(* IEC 61131-3 sources: trust-platform/examples/OSCAT/cip_wash_state/oop/src, 3 files *)

(* ---- Main.st ---- *)
(* Pattern role: ICipState is the contract boundary for the State example. *)
INTERFACE ICipState
    PROPERTY StateId : INT
    GET
    END_GET
    END_PROPERTY

    METHOD OnEnter
    END_METHOD

    METHOD OnExecute : INT
    VAR_INPUT
        StartCommand : BOOL;
        StepComplete : BOOL;
        ConductivityUs : REAL;
        CausticTempC : REAL;
        FlowOk : BOOL;
        EStopHealthy : BOOL;
    END_VAR
    END_METHOD

    METHOD OnExit
    END_METHOD

    METHOD CanAbort : BOOL
    END_METHOD
END_INTERFACE

(* Pattern role: IdleState is a concrete implementation in the State example. *)
FUNCTION_BLOCK IdleState IMPLEMENTS ICipState
VAR
    Entered : BOOL;
END_VAR

METHOD PUBLIC OnEnter
Entered := TRUE;
END_METHOD

METHOD PUBLIC OnExecute : INT
VAR_INPUT
    StartCommand : BOOL;
    StepComplete : BOOL;
    ConductivityUs : REAL;
    CausticTempC : REAL;
    FlowOk : BOOL;
    EStopHealthy : BOOL;
END_VAR
IF NOT EStopHealthy THEN
    OnExecute := INT#90;
ELSIF StartCommand THEN
    OnExecute := INT#10;
ELSE
    OnExecute := INT#0;
END_IF;
END_METHOD

METHOD PUBLIC OnExit
Entered := FALSE;
END_METHOD

METHOD PUBLIC CanAbort : BOOL
CanAbort := TRUE;
END_METHOD

PUBLIC PROPERTY StateId : INT
GET
    StateId := INT#0;
END_GET
END_PROPERTY
END_FUNCTION_BLOCK

(* Pattern role: PreRinseState is a concrete implementation in the State example. *)
FUNCTION_BLOCK PreRinseState IMPLEMENTS ICipState
METHOD PUBLIC OnEnter
END_METHOD

METHOD PUBLIC OnExecute : INT
VAR_INPUT
    StartCommand : BOOL;
    StepComplete : BOOL;
    ConductivityUs : REAL;
    CausticTempC : REAL;
    FlowOk : BOOL;
    EStopHealthy : BOOL;
END_VAR
IF NOT EStopHealthy OR NOT FlowOk THEN
    OnExecute := INT#90;
ELSIF StepComplete THEN
    OnExecute := INT#20;
ELSE
    OnExecute := INT#10;
END_IF;
END_METHOD

METHOD PUBLIC OnExit
END_METHOD

METHOD PUBLIC CanAbort : BOOL
CanAbort := TRUE;
END_METHOD

PUBLIC PROPERTY StateId : INT
GET
    StateId := INT#10;
END_GET
END_PROPERTY
END_FUNCTION_BLOCK

(* Pattern role: CausticWashState is a concrete implementation in the State example. *)
FUNCTION_BLOCK CausticWashState IMPLEMENTS ICipState
METHOD PUBLIC OnEnter
END_METHOD

METHOD PUBLIC OnExecute : INT
VAR_INPUT
    StartCommand : BOOL;
    StepComplete : BOOL;
    ConductivityUs : REAL;
    CausticTempC : REAL;
    FlowOk : BOOL;
    EStopHealthy : BOOL;
END_VAR
IF NOT EStopHealthy OR NOT FlowOk THEN
    OnExecute := INT#90;
ELSIF CausticTempC < REAL#70.0 THEN
    OnExecute := INT#20;
ELSIF StepComplete THEN
    OnExecute := INT#30;
ELSE
    OnExecute := INT#20;
END_IF;
END_METHOD

METHOD PUBLIC OnExit
END_METHOD

METHOD PUBLIC CanAbort : BOOL
CanAbort := TRUE;
END_METHOD

PUBLIC PROPERTY StateId : INT
GET
    StateId := INT#20;
END_GET
END_PROPERTY
END_FUNCTION_BLOCK

(* Pattern role: IntermediateRinseState is a concrete implementation in the State example. *)
FUNCTION_BLOCK IntermediateRinseState IMPLEMENTS ICipState
METHOD PUBLIC OnEnter
END_METHOD

METHOD PUBLIC OnExecute : INT
VAR_INPUT
    StartCommand : BOOL;
    StepComplete : BOOL;
    ConductivityUs : REAL;
    CausticTempC : REAL;
    FlowOk : BOOL;
    EStopHealthy : BOOL;
END_VAR
IF NOT EStopHealthy OR NOT FlowOk THEN
    OnExecute := INT#90;
ELSIF StepComplete THEN
    OnExecute := INT#40;
ELSE
    OnExecute := INT#30;
END_IF;
END_METHOD

METHOD PUBLIC OnExit
END_METHOD

METHOD PUBLIC CanAbort : BOOL
CanAbort := TRUE;
END_METHOD

PUBLIC PROPERTY StateId : INT
GET
    StateId := INT#30;
END_GET
END_PROPERTY
END_FUNCTION_BLOCK

(* Pattern role: AcidWashState is a concrete implementation in the State example. *)
FUNCTION_BLOCK AcidWashState IMPLEMENTS ICipState
METHOD PUBLIC OnEnter
END_METHOD

METHOD PUBLIC OnExecute : INT
VAR_INPUT
    StartCommand : BOOL;
    StepComplete : BOOL;
    ConductivityUs : REAL;
    CausticTempC : REAL;
    FlowOk : BOOL;
    EStopHealthy : BOOL;
END_VAR
IF NOT EStopHealthy OR NOT FlowOk THEN
    OnExecute := INT#90;
ELSIF StepComplete THEN
    OnExecute := INT#50;
ELSE
    OnExecute := INT#40;
END_IF;
END_METHOD

METHOD PUBLIC OnExit
END_METHOD

METHOD PUBLIC CanAbort : BOOL
CanAbort := TRUE;
END_METHOD

PUBLIC PROPERTY StateId : INT
GET
    StateId := INT#40;
END_GET
END_PROPERTY
END_FUNCTION_BLOCK

(* Pattern role: FinalRinseState is a concrete implementation in the State example. *)
FUNCTION_BLOCK FinalRinseState IMPLEMENTS ICipState
METHOD PUBLIC OnEnter
END_METHOD

METHOD PUBLIC OnExecute : INT
VAR_INPUT
    StartCommand : BOOL;
    StepComplete : BOOL;
    ConductivityUs : REAL;
    CausticTempC : REAL;
    FlowOk : BOOL;
    EStopHealthy : BOOL;
END_VAR
IF NOT EStopHealthy OR NOT FlowOk THEN
    OnExecute := INT#90;
ELSIF ConductivityUs < REAL#50.0 THEN
    OnExecute := INT#100;
ELSE
    OnExecute := INT#50;
END_IF;
END_METHOD

METHOD PUBLIC OnExit
END_METHOD

METHOD PUBLIC CanAbort : BOOL
CanAbort := TRUE;
END_METHOD

PUBLIC PROPERTY StateId : INT
GET
    StateId := INT#50;
END_GET
END_PROPERTY
END_FUNCTION_BLOCK

(* Pattern role: DoneState is a concrete implementation in the State example. *)
FUNCTION_BLOCK DoneState IMPLEMENTS ICipState
METHOD PUBLIC OnEnter
END_METHOD

METHOD PUBLIC OnExecute : INT
VAR_INPUT
    StartCommand : BOOL;
    StepComplete : BOOL;
    ConductivityUs : REAL;
    CausticTempC : REAL;
    FlowOk : BOOL;
    EStopHealthy : BOOL;
END_VAR
OnExecute := INT#100;
END_METHOD

METHOD PUBLIC OnExit
END_METHOD

METHOD PUBLIC CanAbort : BOOL
CanAbort := FALSE;
END_METHOD

PUBLIC PROPERTY StateId : INT
GET
    StateId := INT#100;
END_GET
END_PROPERTY
END_FUNCTION_BLOCK

(* Pattern role: AbortState is a concrete implementation in the State example. *)
FUNCTION_BLOCK AbortState IMPLEMENTS ICipState
METHOD PUBLIC OnEnter
END_METHOD

METHOD PUBLIC OnExecute : INT
VAR_INPUT
    StartCommand : BOOL;
    StepComplete : BOOL;
    ConductivityUs : REAL;
    CausticTempC : REAL;
    FlowOk : BOOL;
    EStopHealthy : BOOL;
END_VAR
OnExecute := INT#90;
END_METHOD

METHOD PUBLIC OnExit
END_METHOD

METHOD PUBLIC CanAbort : BOOL
CanAbort := FALSE;
END_METHOD

PUBLIC PROPERTY StateId : INT
GET
    StateId := INT#90;
END_GET
END_PROPERTY
END_FUNCTION_BLOCK

(* Composition role: CipController owns the collaborating objects used by this State example. *)
FUNCTION_BLOCK CipController
VAR
    Idle : IdleState;
    PreRinse : PreRinseState;
    Caustic : CausticWashState;
    Intermediate : IntermediateRinseState;
    Acid : AcidWashState;
    FinalRinse : FinalRinseState;
    CompleteState : DoneState;
    Abort : AbortState;
    Current : ICipState;
    ConductivityFilter : Pt1Filter;
    CycleCounter : DwordCounter;
    CurrentStateIdValue : INT;
    TransitionCountValue : INT;
    AbortedValue : BOOL;
END_VAR

METHOD PUBLIC Initialize
ConductivityFilter.Initialize();
ConductivityFilter.Configure(TimeConstant := T#1s, Gain := REAL#1.0);
CycleCounter.Initialize();
CycleCounter.Configure(StepSize := DWORD#1, MaxValue := DWORD#16#FFFFFFFF);
Current := Idle;
Current.OnEnter();
CurrentStateIdValue := Current.StateId;
TransitionCountValue := INT#0;
AbortedValue := FALSE;
END_METHOD

METHOD PUBLIC ResolveState : ICipState
VAR_INPUT
    NextId : INT;
END_VAR
IF NextId = INT#10 THEN
    ResolveState := PreRinse;
ELSIF NextId = INT#20 THEN
    ResolveState := Caustic;
ELSIF NextId = INT#30 THEN
    ResolveState := Intermediate;
ELSIF NextId = INT#40 THEN
    ResolveState := Acid;
ELSIF NextId = INT#50 THEN
    ResolveState := FinalRinse;
ELSIF NextId = INT#90 THEN
    ResolveState := Abort;
ELSIF NextId = INT#100 THEN
    ResolveState := CompleteState;
ELSE
    ResolveState := Idle;
END_IF;
END_METHOD

METHOD PUBLIC Update : INT
VAR_INPUT
    StartCommand : BOOL;
    StepComplete : BOOL;
    ConductivityUs : REAL;
    CausticTempC : REAL;
    FlowOk : BOOL;
    EStopHealthy : BOOL;
END_VAR
VAR
    NextId : INT;
END_VAR
(* ConductivityFilter is declared and updated for telemetry/HMI use only.
   FinalRinseState compares against the raw ConductivityUs because the
   PT1 filter time constant (1 s) would otherwise delay the wash-complete
   decision past one scan cycle. A production CIP could drive the state
   from the filtered value with a longer minimum-rinse time. *)
ConductivityFilter.Update(Sample := ConductivityUs);
NextId := Current.OnExecute(StartCommand := StartCommand, StepComplete := StepComplete, ConductivityUs := ConductivityUs, CausticTempC := CausticTempC, FlowOk := FlowOk, EStopHealthy := EStopHealthy);
IF NextId <> Current.StateId THEN
    Current.OnExit();
    Current := ResolveState(NextId := NextId);
    Current.OnEnter();
    CurrentStateIdValue := Current.StateId;
    TransitionCountValue := TransitionCountValue + INT#1;
    IF CurrentStateIdValue = INT#90 THEN
        AbortedValue := TRUE;
    ELSIF CurrentStateIdValue = INT#100 THEN
        CycleCounter.Update(Up := TRUE, Down := FALSE);
    END_IF;
END_IF;
Update := CurrentStateIdValue;
END_METHOD

PUBLIC PROPERTY CurrentStateId : INT
GET
    CurrentStateId := CurrentStateIdValue;
END_GET
END_PROPERTY

PUBLIC PROPERTY TransitionCount : INT
GET
    TransitionCount := TransitionCountValue;
END_GET
END_PROPERTY

PUBLIC PROPERTY CycleCount : DWORD
GET
    CycleCount := CycleCounter.Count;
END_GET
END_PROPERTY

PUBLIC PROPERTY Aborted : BOOL
GET
    Aborted := AbortedValue;
END_GET
END_PROPERTY
END_FUNCTION_BLOCK

(* Scan role: Main wires the example objects and exposes the PLC call path under test. *)
PROGRAM Main
VAR
    Cip : CipController;
    Initialized : BOOL;
    StartCommand : BOOL;
    StepComplete : BOOL;
    EStopHealthy : BOOL;
    FlowOk : BOOL;
    ConductivityRaw : INT;
    CausticTempRaw : INT;
    PumpEnableOut : BOOL;
    DrainValveOut : BOOL;
    AlarmOut : BOOL;
END_VAR

(* Initialize once on cold start; scanning Initialize every cycle would
   reset the state machine to Idle and clear retained counters. *)
IF NOT Initialized THEN
    Cip.Initialize();
    Initialized := TRUE;
END_IF;
Cip.Update(StartCommand := StartCommand, StepComplete := StepComplete, ConductivityUs := INT_TO_REAL(ConductivityRaw), CausticTempC := INT_TO_REAL(CausticTempRaw), FlowOk := FlowOk, EStopHealthy := EStopHealthy);
PumpEnableOut := (Cip.CurrentStateId >= INT#10) AND (Cip.CurrentStateId < INT#90);
DrainValveOut := Cip.CurrentStateId = INT#90;
AlarmOut := Cip.Aborted;
END_PROGRAM

(* ---- Configuration.st ---- *)
CONFIGURATION CipWashStateOopConfiguration
RESOURCE Cpu0 ON PLC
    TASK MainTask (INTERVAL := T#100ms, PRIORITY := 1);
    PROGRAM Cip WITH MainTask : Main;
END_RESOURCE
VAR_CONFIG
    Cip.StartCommand AT %IX0.0 : BOOL;
    Cip.StepComplete AT %IX0.1 : BOOL;
    Cip.EStopHealthy AT %IX0.2 : BOOL;
    Cip.FlowOk AT %IX0.3 : BOOL;
    Cip.ConductivityRaw AT %IW0 : INT;
    Cip.CausticTempRaw AT %IW2 : INT;
    Cip.PumpEnableOut AT %QX0.0 : BOOL;
    Cip.DrainValveOut AT %QX0.1 : BOOL;
    Cip.AlarmOut AT %QX0.2 : BOOL;
END_VAR
END_CONFIGURATION

(* ---- Tests.st ---- *)
TEST_PROGRAM CipStateObjectsAdvanceThroughSequence
VAR
    Cip : CipController;
END_VAR

Cip.Initialize();
ASSERT_EQUAL(EXPECTED := INT#10, ACTUAL := Cip.Update(StartCommand := TRUE, StepComplete := FALSE, ConductivityUs := REAL#200.0, CausticTempC := REAL#75.0, FlowOk := TRUE, EStopHealthy := TRUE));
ASSERT_EQUAL(EXPECTED := INT#20, ACTUAL := Cip.Update(StartCommand := FALSE, StepComplete := TRUE, ConductivityUs := REAL#200.0, CausticTempC := REAL#75.0, FlowOk := TRUE, EStopHealthy := TRUE));
ASSERT_EQUAL(EXPECTED := INT#30, ACTUAL := Cip.Update(StartCommand := FALSE, StepComplete := TRUE, ConductivityUs := REAL#200.0, CausticTempC := REAL#75.0, FlowOk := TRUE, EStopHealthy := TRUE));
ASSERT_EQUAL(EXPECTED := INT#40, ACTUAL := Cip.Update(StartCommand := FALSE, StepComplete := TRUE, ConductivityUs := REAL#200.0, CausticTempC := REAL#75.0, FlowOk := TRUE, EStopHealthy := TRUE));
ASSERT_EQUAL(EXPECTED := INT#50, ACTUAL := Cip.Update(StartCommand := FALSE, StepComplete := TRUE, ConductivityUs := REAL#200.0, CausticTempC := REAL#75.0, FlowOk := TRUE, EStopHealthy := TRUE));
ASSERT_EQUAL(EXPECTED := INT#100, ACTUAL := Cip.Update(StartCommand := FALSE, StepComplete := FALSE, ConductivityUs := REAL#20.0, CausticTempC := REAL#75.0, FlowOk := TRUE, EStopHealthy := TRUE));
ASSERT_EQUAL(EXPECTED := DWORD#1, ACTUAL := Cip.CycleCount);
END_TEST_PROGRAM

TEST_PROGRAM CipStateObjectsAbortFromActiveStep
VAR
    Cip : CipController;
END_VAR

Cip.Initialize();
Cip.Update(StartCommand := TRUE, StepComplete := FALSE, ConductivityUs := REAL#200.0, CausticTempC := REAL#75.0, FlowOk := TRUE, EStopHealthy := TRUE);
ASSERT_EQUAL(EXPECTED := INT#90, ACTUAL := Cip.Update(StartCommand := FALSE, StepComplete := FALSE, ConductivityUs := REAL#200.0, CausticTempC := REAL#75.0, FlowOk := FALSE, EStopHealthy := TRUE));
ASSERT_TRUE(IN := Cip.Aborted);
END_TEST_PROGRAM

(* Integration test: simulates the PROGRAM Main scan loop with the
   Init-once guard. Catches the "Initialize every cycle" bug — without
   the guard, the state machine resets to Idle on every iteration and
   never reaches Done. *)
TEST_PROGRAM CipScanLoopWithInitGuardProgressesThroughSequence
VAR
    Cip : CipController;
    Initialized : BOOL;
    I : INT;
    StateValue : INT;
END_VAR

FOR I := 1 TO 6 DO
    IF NOT Initialized THEN
        Cip.Initialize();
        Initialized := TRUE;
    END_IF;
    CASE I OF
        INT#1: StateValue := Cip.Update(StartCommand := TRUE,  StepComplete := FALSE, ConductivityUs := REAL#200.0, CausticTempC := REAL#75.0, FlowOk := TRUE, EStopHealthy := TRUE);
        INT#2: StateValue := Cip.Update(StartCommand := FALSE, StepComplete := TRUE,  ConductivityUs := REAL#200.0, CausticTempC := REAL#75.0, FlowOk := TRUE, EStopHealthy := TRUE);
        INT#3: StateValue := Cip.Update(StartCommand := FALSE, StepComplete := TRUE,  ConductivityUs := REAL#200.0, CausticTempC := REAL#75.0, FlowOk := TRUE, EStopHealthy := TRUE);
        INT#4: StateValue := Cip.Update(StartCommand := FALSE, StepComplete := TRUE,  ConductivityUs := REAL#200.0, CausticTempC := REAL#75.0, FlowOk := TRUE, EStopHealthy := TRUE);
        INT#5: StateValue := Cip.Update(StartCommand := FALSE, StepComplete := TRUE,  ConductivityUs := REAL#200.0, CausticTempC := REAL#75.0, FlowOk := TRUE, EStopHealthy := TRUE);
        INT#6: StateValue := Cip.Update(StartCommand := FALSE, StepComplete := FALSE, ConductivityUs := REAL#20.0,  CausticTempC := REAL#75.0, FlowOk := TRUE, EStopHealthy := TRUE);
    END_CASE;
END_FOR;
ASSERT_EQUAL(EXPECTED := INT#100, ACTUAL := StateValue);
ASSERT_EQUAL(EXPECTED := DWORD#1, ACTUAL := Cip.CycleCount);
END_TEST_PROGRAM

(* Anti-pattern test: explicitly demonstrates that calling Initialize on
   every cycle resets the state machine. If a future change removes the
   Init-once guard from Main, this test pins the contract: re-init each
   cycle cannot reach the wash-complete state. *)
TEST_PROGRAM CipReinitializingEveryCycleResetsStateMachine
VAR
    Cip : CipController;
    I : INT;
    StateValue : INT;
END_VAR

FOR I := 1 TO 6 DO
    Cip.Initialize();
    StateValue := Cip.Update(StartCommand := TRUE, StepComplete := TRUE, ConductivityUs := REAL#20.0, CausticTempC := REAL#75.0, FlowOk := TRUE, EStopHealthy := TRUE);
END_FOR;
(* Re-initializing every cycle: state machine cannot get past PreRinse *)
ASSERT_TRUE(IN := StateValue <= INT#10);
ASSERT_EQUAL(EXPECTED := DWORD#0, ACTUAL := Cip.CycleCount);
END_TEST_PROGRAM

(* Idle state edge cases: e-stop loss aborts before start; no command holds at 0. *)
TEST_PROGRAM CipIdleStateBranchesCovered
VAR
    Cip : CipController;
END_VAR
Cip.Initialize();
(* No start command: state stays at 0 *)
ASSERT_EQUAL(EXPECTED := INT#0, ACTUAL := Cip.Update(StartCommand := FALSE, StepComplete := FALSE, ConductivityUs := REAL#200.0, CausticTempC := REAL#75.0, FlowOk := TRUE, EStopHealthy := TRUE));
(* E-stop loss while idle: state goes to abort (90) *)
ASSERT_EQUAL(EXPECTED := INT#90, ACTUAL := Cip.Update(StartCommand := TRUE, StepComplete := FALSE, ConductivityUs := REAL#200.0, CausticTempC := REAL#75.0, FlowOk := TRUE, EStopHealthy := FALSE));
ASSERT_TRUE(IN := Cip.Aborted);
END_TEST_PROGRAM

(* CausticWash temperature gate: must reach 70 C before stepping forward. *)
TEST_PROGRAM CipCausticWashHoldsBelowTemperatureThreshold
VAR
    Cip : CipController;
END_VAR
Cip.Initialize();
(* Drive into caustic wash *)
Cip.Update(StartCommand := TRUE, StepComplete := FALSE, ConductivityUs := REAL#200.0, CausticTempC := REAL#75.0, FlowOk := TRUE, EStopHealthy := TRUE);
Cip.Update(StartCommand := FALSE, StepComplete := TRUE, ConductivityUs := REAL#200.0, CausticTempC := REAL#75.0, FlowOk := TRUE, EStopHealthy := TRUE);
ASSERT_EQUAL(EXPECTED := INT#20, ACTUAL := Cip.CurrentStateId);
(* Below threshold even with StepComplete - stays in caustic *)
ASSERT_EQUAL(EXPECTED := INT#20, ACTUAL := Cip.Update(StartCommand := FALSE, StepComplete := TRUE, ConductivityUs := REAL#200.0, CausticTempC := REAL#69.9, FlowOk := TRUE, EStopHealthy := TRUE));
(* Below 70 without StepComplete - stays *)
ASSERT_EQUAL(EXPECTED := INT#20, ACTUAL := Cip.Update(StartCommand := FALSE, StepComplete := FALSE, ConductivityUs := REAL#200.0, CausticTempC := REAL#65.0, FlowOk := TRUE, EStopHealthy := TRUE));
(* At 70 + StepComplete - advances to intermediate rinse (30) *)
ASSERT_EQUAL(EXPECTED := INT#30, ACTUAL := Cip.Update(StartCommand := FALSE, StepComplete := TRUE, ConductivityUs := REAL#200.0, CausticTempC := REAL#70.0, FlowOk := TRUE, EStopHealthy := TRUE));
END_TEST_PROGRAM

(* FinalRinse conductivity gate: must drop below 50 uS/cm to complete. *)
TEST_PROGRAM CipFinalRinseHoldsAboveConductivityThreshold
VAR
    Cip : CipController;
END_VAR
Cip.Initialize();
(* Drive through to FinalRinse *)
Cip.Update(StartCommand := TRUE, StepComplete := FALSE, ConductivityUs := REAL#200.0, CausticTempC := REAL#75.0, FlowOk := TRUE, EStopHealthy := TRUE);
Cip.Update(StartCommand := FALSE, StepComplete := TRUE, ConductivityUs := REAL#200.0, CausticTempC := REAL#75.0, FlowOk := TRUE, EStopHealthy := TRUE);
Cip.Update(StartCommand := FALSE, StepComplete := TRUE, ConductivityUs := REAL#200.0, CausticTempC := REAL#75.0, FlowOk := TRUE, EStopHealthy := TRUE);
Cip.Update(StartCommand := FALSE, StepComplete := TRUE, ConductivityUs := REAL#200.0, CausticTempC := REAL#75.0, FlowOk := TRUE, EStopHealthy := TRUE);
Cip.Update(StartCommand := FALSE, StepComplete := TRUE, ConductivityUs := REAL#200.0, CausticTempC := REAL#75.0, FlowOk := TRUE, EStopHealthy := TRUE);
ASSERT_EQUAL(EXPECTED := INT#50, ACTUAL := Cip.CurrentStateId);
(* Conductivity above 50: stays in FinalRinse *)
ASSERT_EQUAL(EXPECTED := INT#50, ACTUAL := Cip.Update(StartCommand := FALSE, StepComplete := FALSE, ConductivityUs := REAL#100.0, CausticTempC := REAL#75.0, FlowOk := TRUE, EStopHealthy := TRUE));
(* Just at 50: stays (strict less-than required) *)
ASSERT_EQUAL(EXPECTED := INT#50, ACTUAL := Cip.Update(StartCommand := FALSE, StepComplete := FALSE, ConductivityUs := REAL#50.0, CausticTempC := REAL#75.0, FlowOk := TRUE, EStopHealthy := TRUE));
(* Just below 50: completes *)
ASSERT_EQUAL(EXPECTED := INT#100, ACTUAL := Cip.Update(StartCommand := FALSE, StepComplete := FALSE, ConductivityUs := REAL#49.9, CausticTempC := REAL#75.0, FlowOk := TRUE, EStopHealthy := TRUE));
END_TEST_PROGRAM

(* Done state is terminal: any further Update returns 100. *)
TEST_PROGRAM CipDoneStateIsTerminal
VAR
    Cip : CipController;
END_VAR
Cip.Initialize();
(* Drive to done *)
Cip.Update(StartCommand := TRUE, StepComplete := FALSE, ConductivityUs := REAL#200.0, CausticTempC := REAL#75.0, FlowOk := TRUE, EStopHealthy := TRUE);
Cip.Update(StartCommand := FALSE, StepComplete := TRUE, ConductivityUs := REAL#200.0, CausticTempC := REAL#75.0, FlowOk := TRUE, EStopHealthy := TRUE);
Cip.Update(StartCommand := FALSE, StepComplete := TRUE, ConductivityUs := REAL#200.0, CausticTempC := REAL#75.0, FlowOk := TRUE, EStopHealthy := TRUE);
Cip.Update(StartCommand := FALSE, StepComplete := TRUE, ConductivityUs := REAL#200.0, CausticTempC := REAL#75.0, FlowOk := TRUE, EStopHealthy := TRUE);
Cip.Update(StartCommand := FALSE, StepComplete := TRUE, ConductivityUs := REAL#200.0, CausticTempC := REAL#75.0, FlowOk := TRUE, EStopHealthy := TRUE);
Cip.Update(StartCommand := FALSE, StepComplete := FALSE, ConductivityUs := REAL#20.0, CausticTempC := REAL#75.0, FlowOk := TRUE, EStopHealthy := TRUE);
ASSERT_EQUAL(EXPECTED := INT#100, ACTUAL := Cip.CurrentStateId);
(* Subsequent Updates with any inputs keep state at 100 *)
ASSERT_EQUAL(EXPECTED := INT#100, ACTUAL := Cip.Update(StartCommand := TRUE, StepComplete := TRUE, ConductivityUs := REAL#5.0, CausticTempC := REAL#80.0, FlowOk := TRUE, EStopHealthy := TRUE));
ASSERT_EQUAL(EXPECTED := INT#100, ACTUAL := Cip.Update(StartCommand := FALSE, StepComplete := FALSE, ConductivityUs := REAL#200.0, CausticTempC := REAL#0.0, FlowOk := FALSE, EStopHealthy := FALSE));
END_TEST_PROGRAM

(* Abort state is terminal: any further Update returns 90 even with all inputs healthy. *)
TEST_PROGRAM CipAbortStateIsTerminal
VAR
    Cip : CipController;
END_VAR
Cip.Initialize();
Cip.Update(StartCommand := TRUE, StepComplete := FALSE, ConductivityUs := REAL#200.0, CausticTempC := REAL#75.0, FlowOk := TRUE, EStopHealthy := TRUE);
Cip.Update(StartCommand := FALSE, StepComplete := FALSE, ConductivityUs := REAL#200.0, CausticTempC := REAL#75.0, FlowOk := FALSE, EStopHealthy := TRUE);
ASSERT_EQUAL(EXPECTED := INT#90, ACTUAL := Cip.CurrentStateId);
(* Healthy inputs after abort: still at 90 *)
ASSERT_EQUAL(EXPECTED := INT#90, ACTUAL := Cip.Update(StartCommand := TRUE, StepComplete := TRUE, ConductivityUs := REAL#20.0, CausticTempC := REAL#75.0, FlowOk := TRUE, EStopHealthy := TRUE));
ASSERT_TRUE(IN := Cip.Aborted);
END_TEST_PROGRAM

(* CycleCount increments only on Done transitions, not on Abort. *)
TEST_PROGRAM CipCycleCountTracksOnlyCompletions
VAR
    Cip : CipController;
END_VAR
Cip.Initialize();
(* First wash: complete cycle - cycle count := 1 *)
Cip.Update(StartCommand := TRUE, StepComplete := FALSE, ConductivityUs := REAL#200.0, CausticTempC := REAL#75.0, FlowOk := TRUE, EStopHealthy := TRUE);
Cip.Update(StartCommand := FALSE, StepComplete := TRUE, ConductivityUs := REAL#200.0, CausticTempC := REAL#75.0, FlowOk := TRUE, EStopHealthy := TRUE);
Cip.Update(StartCommand := FALSE, StepComplete := TRUE, ConductivityUs := REAL#200.0, CausticTempC := REAL#75.0, FlowOk := TRUE, EStopHealthy := TRUE);
Cip.Update(StartCommand := FALSE, StepComplete := TRUE, ConductivityUs := REAL#200.0, CausticTempC := REAL#75.0, FlowOk := TRUE, EStopHealthy := TRUE);
Cip.Update(StartCommand := FALSE, StepComplete := TRUE, ConductivityUs := REAL#200.0, CausticTempC := REAL#75.0, FlowOk := TRUE, EStopHealthy := TRUE);
Cip.Update(StartCommand := FALSE, StepComplete := FALSE, ConductivityUs := REAL#20.0, CausticTempC := REAL#75.0, FlowOk := TRUE, EStopHealthy := TRUE);
ASSERT_EQUAL(EXPECTED := DWORD#1, ACTUAL := Cip.CycleCount);

(* Second wash starts after Done is terminal - CycleCount unchanged *)
Cip.Update(StartCommand := TRUE, StepComplete := TRUE, ConductivityUs := REAL#20.0, CausticTempC := REAL#75.0, FlowOk := TRUE, EStopHealthy := TRUE);
ASSERT_EQUAL(EXPECTED := DWORD#1, ACTUAL := Cip.CycleCount);
END_TEST_PROGRAM

(* PreRinse and IntermediateRinse: flow loss aborts at any moment. *)
TEST_PROGRAM CipFlowLossAbortsRinseStates
VAR
    Cip : CipController;
END_VAR
Cip.Initialize();
(* Enter PreRinse, lose flow *)
Cip.Update(StartCommand := TRUE, StepComplete := FALSE, ConductivityUs := REAL#200.0, CausticTempC := REAL#75.0, FlowOk := TRUE, EStopHealthy := TRUE);
ASSERT_EQUAL(EXPECTED := INT#90, ACTUAL := Cip.Update(StartCommand := FALSE, StepComplete := FALSE, ConductivityUs := REAL#200.0, CausticTempC := REAL#75.0, FlowOk := FALSE, EStopHealthy := TRUE));
ASSERT_TRUE(IN := Cip.Aborted);
END_TEST_PROGRAM

(* AcidWash flow loss aborts. *)
TEST_PROGRAM CipFlowLossAbortsAcidWash
VAR
    Cip : CipController;
END_VAR
Cip.Initialize();
(* Drive to AcidWash *)
Cip.Update(StartCommand := TRUE, StepComplete := FALSE, ConductivityUs := REAL#200.0, CausticTempC := REAL#75.0, FlowOk := TRUE, EStopHealthy := TRUE);
Cip.Update(StartCommand := FALSE, StepComplete := TRUE, ConductivityUs := REAL#200.0, CausticTempC := REAL#75.0, FlowOk := TRUE, EStopHealthy := TRUE);
Cip.Update(StartCommand := FALSE, StepComplete := TRUE, ConductivityUs := REAL#200.0, CausticTempC := REAL#75.0, FlowOk := TRUE, EStopHealthy := TRUE);
Cip.Update(StartCommand := FALSE, StepComplete := TRUE, ConductivityUs := REAL#200.0, CausticTempC := REAL#75.0, FlowOk := TRUE, EStopHealthy := TRUE);
ASSERT_EQUAL(EXPECTED := INT#40, ACTUAL := Cip.CurrentStateId);
(* Flow loss while in AcidWash *)
ASSERT_EQUAL(EXPECTED := INT#90, ACTUAL := Cip.Update(StartCommand := FALSE, StepComplete := FALSE, ConductivityUs := REAL#200.0, CausticTempC := REAL#75.0, FlowOk := FALSE, EStopHealthy := TRUE));
END_TEST_PROGRAM

(* TransitionCount accumulates exactly one increment per state change. *)
TEST_PROGRAM CipTransitionCountMatchesStateChanges
VAR
    Cip : CipController;
END_VAR
Cip.Initialize();
(* Each StepComplete = one transition *)
Cip.Update(StartCommand := TRUE, StepComplete := FALSE, ConductivityUs := REAL#200.0, CausticTempC := REAL#75.0, FlowOk := TRUE, EStopHealthy := TRUE);
ASSERT_EQUAL(EXPECTED := INT#1, ACTUAL := Cip.TransitionCount);
(* Stay in PreRinse - no transition *)
Cip.Update(StartCommand := FALSE, StepComplete := FALSE, ConductivityUs := REAL#200.0, CausticTempC := REAL#75.0, FlowOk := TRUE, EStopHealthy := TRUE);
ASSERT_EQUAL(EXPECTED := INT#1, ACTUAL := Cip.TransitionCount);
(* Step complete - transit to caustic *)
Cip.Update(StartCommand := FALSE, StepComplete := TRUE, ConductivityUs := REAL#200.0, CausticTempC := REAL#75.0, FlowOk := TRUE, EStopHealthy := TRUE);
ASSERT_EQUAL(EXPECTED := INT#2, ACTUAL := Cip.TransitionCount);
END_TEST_PROGRAM
